Fanuc KAREL source: KD00027.KL

PROGRAM KD00027
%NOLOCKGROUP
VAR
  I: INTEGER
  J: INTEGER
  B: BOOLEAN
  R: REAL
  S: STRING[80]
BEGIN
  CONDITION[1]:
  WHEN EVENT[1] DO
    I = 1
  ENDCONDITION
END KD00027
